Staubli VAL3: actCmd.pjx

--- actCmd.pjx ---
Parameters version=s8.10.2Cs9_BS1991 stackSize=5000 millimeterUnit=true
Data file=actCmd.dtx

--- actCmd.dtx ---
public num nMoveID
public num nActionID
public bool bActFinish
public string sActName
